(* IEC 61131-3 sources: plc-vscode/tests/st/all/trust-platform/crates/trust-runtime/tests/fixtures/opcua/program, 1 file *)

(* ---- main.st ---- *)
CONFIGURATION OpcUaFixture
VAR_GLOBAL
    counter : DINT := 42;
    ready : BOOL := TRUE;
    name : STRING := 'pump';
END_VAR
TASK Fast (INTERVAL := T#10ms, PRIORITY := 0);
PROGRAM App WITH Fast : Main;
END_CONFIGURATION

PROGRAM Main
END_PROGRAM
